// TIA Portal project "AT4B_Start" (V18)

(* hardware
DEVICE "PLC_1_Station"  S7-1500 station
   slot 0: "Profilschiene_0"  Rack  6ES7 590-1***0-0AA0
   slot 1: "PLC_1"  CPU 1516-3 PN/DP  6ES7 516-3AN02-0AB0  V2.8
      slot 3: "CPU-Display_1"  6ES7591-1BA00-0AA0
      slot 32768: "PROFINET-Schnittstelle_1"  X1
         slot 32769: "Port_1"  X1 P1
         slot 32770: "Port_2"  X1 P2
      slot 33024: "PROFINET-Schnittstelle_2"  X2
         slot 33025: "Port_1"  X2 P1
      slot 33280: "DP-Schnittstelle_1"  X3
      slot 34817: "Virtual CP interface port_1"  Virtual CP interface port  Virtual CP interface port
DEVICE "HMI_1"  KTP1200 Basic DP
   slot 0: "HMI_1"  KTP1200 Basic DP  6AV2 123-2MA03-0AX0  15.1.0.0
   slot 1: "HMI_RT_1"  KTP1200 Basic DP  6AV2 123-2MA03-0AX0  15.1.0.0
   slot 7: "HMI_1.MPI/DP_CP_1"  MPI/DP Interface  15.0.1.0
DEVICE "HMI_2"  KTP1200 Basic PN
   slot 0: "HMI_2"  KTP1200 Basic PN  6AV2 123-2MB03-0AX0  17.0.0.0
   slot 1: "HMI_RT_2"  KTP1200 Basic PN  6AV2 123-2MB03-0AX0  17.0.0.0
   slot 5: "HMI_2.IE_CP_1"  PROFINET Interface  17.0.0.0
      slot 1: "PROFINET Schnittstelle_1"  PROFINET Interface
         slot 1: "Port_1"  Port
*)

// ===== PLC "PLC_1"  CPU 1516-3 PN/DP =====

VAR_GLOBAL   // PLC tag table "Private_Linktest"
   "ProofInput1" AT %M2.0 : LReal;
   "ProofInput2" AT %M10.0 : LReal;
   "ProofOutput" AT %M18.0 : LReal;
   "ProofFlag" AT %M0.0 : Bool;
END_VAR

ORGANIZATION_BLOCK "Main"   // OB1, FBD, ProgramCycle
TITLE = "Main Program Sweep (Cycle)"
{ S7_Optimized_Access := 'TRUE' }
VERSION : 0.1
   VAR_INPUT
      Initial_Call : Bool;   // Initial call of this OB
      Remanence : Bool;   // =True, if remanent data are available
   END_VAR
BEGIN
END_ORGANIZATION_BLOCK

(* ===== HMI "HMI_RT_1" =====
connection "HMI_Verbindung_1": IF1 B, SMART_S7_1500_OMS
connection "HMI_Verbindung_3": IF1 B, SMART_S7_1500_OMS
connection "Verbindung_1": IF1 B, SMART_S7_1500_OMS

HMI tags "Private_Linktest"
   "ProofInput1" : LReal AT %M2.0, 1 s
   "ProofInput2" : LReal AT %M10.0, 1 s
   "ProofOutput" : LReal AT %M18.0, 1 s
   "ProofFlag" : Bool AT %M0.0, 1 s

screen "Verbindungspruefung" 1280x800
   IOField "Linktest_ProofInput1" at 64,120 size 1152x76; HelpText 'Private Kopplungspruefung, keine Rechenfunktion. Testwert eingeben und mit Enter bestaetigen.'; FormatPattern s999999999.999; Unit Eingabe 1 | M2.0 | HMI -> SPS
      ProcessValue <- "ProofInput1"
   IOField "Linktest_ProofInput2" at 64,300 size 1152x76; HelpText 'Private Kopplungspruefung, keine Rechenfunktion. Testwert eingeben und mit Enter bestaetigen.'; FormatPattern s999999999.999; Unit Eingabe 2 | M10.0 | HMI -> SPS
      ProcessValue <- "ProofInput2"
   IOField "Linktest_ProofOutput" at 64,480 size 1152x76; HelpText 'Private Kopplungspruefung, keine Rechenfunktion. Nur Anzeige des SPS-Merkers.'; FormatPattern s999999999.999; Unit Ausgabe | M18.0 | SPS -> HMI
      ProcessValue <- "ProofOutput"
*)

(* ===== HMI "HMI_RT_2" =====
connection "HMI_Verbindung_2": ETHERNET, SMART_S7_1500_OMS
connection "Pruefung_X1": ETHERNET, SMART_S7_1500_OMS

HMI tags "Private_Linktest"
   "ProofInput1" : LReal AT %M2.0, 1 s
   "ProofInput2" : LReal AT %M10.0, 1 s
   "ProofOutput" : LReal AT %M18.0, 1 s
   "ProofFlag" : Bool AT %M0.0, 1 s
   "InternalCheck" : LReal, internal
   "NativeProbe" : LReal AT %M18.0, 1 s

screen "Verbindungspruefung" 1280x800
   IOField "Linktest_ProofInput1" at 64,120 size 1152x76; HelpText 'Private Kopplungspruefung, keine Rechenfunktion. Testwert eingeben und mit Enter bestaetigen.'; FormatPattern s999999999.999; Unit Eingabe 1 | M2.0 | HMI -> SPS
      ProcessValue <- "ProofInput1"
   IOField "Linktest_ProofInput2" at 64,300 size 1152x76; HelpText 'Private Kopplungspruefung, keine Rechenfunktion. Testwert eingeben und mit Enter bestaetigen.'; FormatPattern s999999999.999; Unit Eingabe 2 | M10.0 | HMI -> SPS
      ProcessValue <- "ProofInput2"
   IOField "Linktest_ProofOutput" at 64,480 size 1152x76; HelpText 'Private Kopplungspruefung, keine Rechenfunktion. Nur Anzeige des SPS-Merkers.'; FormatPattern s999999999.999; Unit Ausgabe | M18.0 | SPS -> HMI
      ProcessValue <- "ProofOutput"
   AlarmView "Meldeanzeige_1" at 0,0 size 600x300
*)